SUBAPPLICATION RedWhiteBackground3SC (* Hintergrundfarbe (TRUE -> Rot, FALSE -> Weiß) für 3 Objekte (Kompakt) *)
  (* Standard: 61499-2 *)
  (* Version 1.0, 2026-07-21, franz, Meisterschulen am Ostbahnhof *)
  PACKAGE MyLib::sys;
  IMPORT isobus::UT::Q::types::s2ObjectIDs;
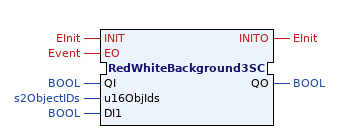
  EVENT_INPUT
    INIT : EInit; (* Initialization Request *)
    EO;
  END_EVENT
  EVENT_OUTPUT
    INITO : EInit; (* Initialization Confirm *)
  END_EVENT
  VAR_INPUT
    QI : BOOL := TRUE; (* Quality Input - TRUE to enable service *)
    u16ObjIds : isobus::UT::Q::types::s2ObjectIDs;
    DI1 : BOOL; (* Selector *)
  END_VAR
  VAR_OUTPUT
    QO : BOOL; (* Quality Output - TRUE if service executed successfully *)
  END_VAR
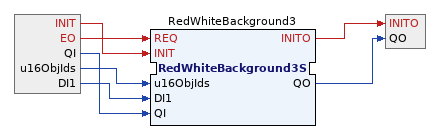
  SUBAPPS
    RedWhiteBackground3 : MyLib::sys::RedWhiteBackground3S;
  END_SUBAPPS
  EVENT_CONNECTIONS
    EO TO RedWhiteBackground3.REQ;
    INIT TO RedWhiteBackground3.INIT;
    RedWhiteBackground3.INITO TO INITO;
  END_CONNECTIONS
  DATA_CONNECTIONS
    u16ObjIds TO RedWhiteBackground3.u16ObjIds;
    DI1 TO RedWhiteBackground3.DI1;
    QI TO RedWhiteBackground3.QI;
    RedWhiteBackground3.QO TO QO;
  END_CONNECTIONS
END_SUBAPPLICATION
